{attribute 'qualified_only' := ''}
{attribute 'strict' := ''}
TYPE E_MCAxisStates :
(
	MC_AXISSTATE_UNDEFINED,
	MC_AXISSTATE_DISABLED,
	MC_AXISSTATE_STANDSTILL,
	MC_AXISSTATE_ERRORSTOP,
	MC_AXISSTATE_STOPPING,
	MC_AXISSTATE_HOMING,
	MC_AXISSTATE_DISCRETEMOTION,
	MC_AXISSTATE_CONTINOUSMOTION,
	MC_AXISSTATE_SYNCHRONIZEDMOTION
);
END_TYPE

(* stored: Version 1.1.0.1, ProductVersion 3.1.4024.12
   DUT E_MCAxisStates: Id {86800532-441f-4161-a371-3d9561ab4c70} *)
